(* IEC 61131-3 sources: JingjiangArm/moonboxpro_arm_8.4/Application/Application/数据类型/通讯协议/云影/读写内容/附属内容, 7 files *)

(* ---- StWrRd_AxisCfg.st ---- *)
(*@CES
Name=StWrRd_AxisCfg
Type=Gvl
TypeGuid=2db5746d-d284-4425-9f7f-2663a34b0ebc
Guid=0dd870ae-2077-401c-9916-294cbac50220
HasDeclaration=True
HasImplementation=False
*)
{DECLARATION}
{attribute 'pack_mode' := '1'}//系统配置
TYPE StWrRd_AxisCfg :
STRUCT
	xAxisProf_Enable: BIT;(*轴打开*)
	xAxisProf_MotRev: BIT;(*运动反向*)
	xAxisProf_SamRev: BIT;(*采样方向*)
	xAxisProf_Rsv1: BIT;(*预留*)
	xAxisProf_Rsv2: BIT;(*预留*)
	xAxisProf_Rsv3: BIT;(*预留*)
	xAxisProf_Rsv4: BIT;(*预留*)
	xAxisProf_Rsv5: BIT;(*预留*)

	//2025.11.1.104728两个字节作为站号通讯
	iSid: INT;
//	abyRsv: ARRAY [1..2] OF BYTE;(*预留两个字节方便增加其他内容*)
END_STRUCT
END_TYPE

{IMPLEMENTATION}

(* ---- StWrRd_MechanicalType.st ---- *)
(*@CES
Name=StWrRd_MechanicalType
Type=Gvl
TypeGuid=2db5746d-d284-4425-9f7f-2663a34b0ebc
Guid=03e174c8-9f43-4388-8870-9d21820ee6bb
HasDeclaration=True
HasImplementation=False
*)
{DECLARATION}
{attribute 'pack_mode' := '1'}
TYPE StWrRd_MechanicalType :
STRUCT
	byMachanicalTypeId: BYTE;(*1摆臂2直压3PVC直压4等料长5力达欧诺直压*)
	abyrsv: ARRAY [1..19] OF BYTE;//先放19个字节在这里放其他预套准相关内容|例如按钮
	abyBuffMechanicalParam: ARRAY [1..200] OF BYTE;(*机械参数*)
	//预留200字节用于通讯机械参数，
		//根据byMachanicalTypeId变量切换通讯内容
		//StMechanicalParam_01/
		//StMechanicalParam_02/
		//StMechanicalParam_03/
		//StMechanicalParam_05
END_STRUCT
END_TYPE

{IMPLEMENTATION}

(* ---- StWrRd_Switch_Grp.st ---- *)
(*@CES
Name=StWrRd_Switch_Grp
Type=Gvl
TypeGuid=2db5746d-d284-4425-9f7f-2663a34b0ebc
Guid=4a26eb77-6c13-4193-b710-63a532b0c18f
HasDeclaration=True
HasImplementation=False
*)
{DECLARATION}
{attribute 'pack_mode' := '1'}//总22字节
TYPE StWrRd_Switch_Grp :
STRUCT
	xSwitch_MachineRev							: BIT;(*反向走料开关*)
	xSwitch_6Inch_Rw							: BIT;(*收料3/6吋选择开关*)
	xSwitch_StartUp								: BIT;(*一键开机开关*)
	xSwitch_DiamMeasureAuto						: BIT;(*自动卷径开关*)
	xSwitch_RollOver							: BIT;(*设备翻料架开关*)
	xSwitch_Thickness							: BIT;(*料膜厚度手自动获取开关*)
	xSwitch_CutDneResetPidEn_Uw					: BIT;(*放料裁切后系数手自动*)
	xSwitch_CutDneResetPidEn_Rw					: BIT;(*收料裁切后系数手自动*)
	xSwitch_AutomaticCutEn_Uw					: BIT;(*放料自动接料是能*)
	xSwitch_AutomaticCutEn_Rw					: BIT;(*放料自动接料是能*)
	xSwitch_AutoAdjust_V_Grp					: BIT;(*整机纵向自动调整开关*)
	xSwitch_AutoAdjust_H_Grp					: BIT;(*整机纵向自动调整开关*)
	xSwitch_Follow_1U_V_Grp						: BIT;(*纵向跟1色开关*)
	xSwitch_Follow_1U_H_Grp						: BIT;(*横向跟1色开关*)
	xSwitch_DiamAuto_Pot						: BIT;(*卷径检测使用电位器*)
	xSwitch_DiamAuto_Enc						: BIT;(*卷径检测使用编码器*)
	xSwitch_DiamAuto_Ultrasonic_S				: BIT;(*卷径检测使用单超声波*)
	xSwitch_DiamAuto_Ultrasonic_D				: BIT;(*卷径检测使用双超声波*)
	xSwitch_DiamAuto_DualParam					: BIT;(*卷径检测双轴参数分开*)
	xSwitch_DebugMode							: BIT;(*调试模式开关*)
	xSwitch_Debug_DiamMeasure_Uw				: BIT;(*放料卷径检测电位器调试开关*)
	xBtn_Diameasure_Confirm_1					: BIT;(*自动卷径标定——1*)
	xBtn_Diameasure_Confirm_2					: BIT;(*自动卷径标定——2*)
	xBtn_Diameasure_Confirm_3					: BIT;(*自动卷径标定——3*)
	xBtn_Diameasure_Confirm_4					: BIT;(*自动卷径标定——4*)
(*2025.11.3.153321收放料绝对值编码器定位等相关开关
原总共42BIT位||重新整理一部分||总共需要14BIT位剩余作为预留*)
	xSwitch_UseAbsEnc_Uw						: BIT;(*放料使用绝对值编码器开关*)
	xSwitch_AxisLocaltion_DualParam_Uw			: BIT;(*放料绝对值编码器定位双轴参数开关*)
	xSwitch_Debug_Axis_Uw						: BIT;(*放料轴运行调试模式*)
	xSwitch_Debug_Uw_CutUpChoose				: BIT;(*放料绝对值编码器定位调试-上下裁选择||TRUE：上裁FALSE：下裁*)
	xSwitch_Debug_Uw_AxisA_Choose				: BIT;(*放料绝对值编码器定位调试-AB轴选择|TRUE:A轴；FALSE:B轴*)
	xBtn_Debug_Uw_Wr							: BIT;(*放料轴定位写入*)
	xBtn_Debug_Uw_MinDiam_Wr					: BIT;(*放料最小径写入*)
	xSwitch_UseAbsEnc_Rw						: BIT;(*收料使用绝对值编码器开关*)
	xSwitch_AxisLocaltion_DualParam_Rw			: BIT;(*收料绝对值编码器定位双轴参数开关*)
	xSwitch_Debug_Axis_Rw						: BIT;(*收料轴运行调试模式*)
	xSwitch_Debug_Rw_CutUpChoose				: BIT;(*收料绝对值编码器定位调试-上下裁选择||TRUE：上裁FALSE：下裁*)
	xSwitch_Debug_Rw_AxisA_Choose				: BIT;(*收料绝对值编码器定位调试-AB轴选择|TRUE:A轴；FALSE:B轴*)
	xSwitch_Debug_Rw_Inch3_CutUpChoose			: BIT;(*收料绝对值编码器定位调试-3/6吋选择|TRUE:3吋；FALSE:6吋*)
	xBtn_Debug_Rw_Wr							: BIT;(*收料轴定位写入*)
//2026.4.25.140018合并结构体|niu.j|增加5个变量
	xSwitch_StartAutoFind	: BIT;(*全自动套印开关*)
	xSwitch_EnFastPress		: BIT;(*当前色找到就合压使能*)
	xSwitch_SaveRS2File		: BIT;(*粗采样保存*)
	xSwitch_RFailure		: BIT;(*全自动套印粗采样失败校准*)
	xSwitch_FFailure		: BIT;(*全自动套印精采样失败校准按钮*)
// 	xRsv_Grp_1									: BIT;
// 	xRsv_Grp_2									: BIT;
// 	xRsv_Grp_3									: BIT;
// 	xRsv_Grp_4									: BIT;
// 	xRsv_Grp_5									: BIT;
//2026.4.25.140311增加结束
	xRsv_Grp_6									: BIT;
	xRsv_Grp_7									: BIT;
	xRsv_Grp_8									: BIT;
	xRsv_Grp_9									: BIT;
	xRsv_Grp_10									: BIT;
	xRsv_Grp_11									: BIT;
	xRsv_Grp_12									: BIT;
	xRsv_Grp_13									: BIT;
	xRsv_Grp_14									: BIT;
	xRsv_Grp_15									: BIT;
	xRsv_Grp_16									: BIT;
	xRsv_Grp_17									: BIT;
	xRsv_Grp_18									: BIT;
//2026.4.28.104338增加异站虚拟码盘重新配置开关xRsv_Grp_19
//	xRsv_Grp_19									: BIT;
	xSwitch_ReSetEncCfg							: BIT;

//bit20和bit21替换为换卷完成放料和收料
// 	xRsv_Grp_20									: BIT;
// 	xRsv_Grp_21									: BIT;
	xBtn_ChangeFilmDn_Uw						: BIT;
	xBtn_ChangeFilmDn_Rw						: BIT;
//2026.04.10.180829结束
//2026.03.11.100402 | + | 使用Bit22作为压力电机自动合压开关
	xSwitch_PressureAuto_Up_Dn							: BIT;
	//xRsv_Grp_22									: BIT;
//2026.2.25.094558 | + | 使用Bit23作为天枢数据保存的开关
	xSwitch_SaveData_GNS						: BIT;
	//xRsv_Grp_23									: BIT;
//2026.02.01.112053 | + | 使用Bit24作为停机维持使能的开关
	xSwitch_KeepServoOn							: BIT;
	//xRsv_Grp_24									: BIT;
//2026.01.27.093334 | + | 使用Bit25和Bit26作为清除报警按钮和回零位的操作标志
	xSwitch_ClearSysAlarm						: BIT;
	xSwitch_BackToHome							: BIT;
// 	xRsv_Grp_25									: BIT;
// 	xRsv_Grp_26									: BIT;
//2026.1.5.151405增加用Bit27和bit28作为收牵压力传感器调整开关和带长调整基准（标准带长/首色带长）开关（暂时只有秦华用）
	xSwitch_TensionAdjust_QH					: BIT;
	xSwitch_PrnLenAdj_Follow_QH					: BIT;
//	xRsv_Grp_27									: BIT;
//	xRsv_Grp_28									: BIT;
(*
	xSwitch_UseAbsEnc_Uw						: BIT;(*放料使用绝对值编码器开关*)
	xSwitch_AxisLocaltion_DualParam_Uw			: BIT;(*放料绝对值编码器定位双轴参数开关*)
	xSwitch_Debug_Axis_Uw						: BIT;(*放料轴运行调试模式*)
	xSwitch_Debug_Uw_CutUpChoose				: BIT;(*放料绝对值编码器定位调试-上裁选择*)
	xSwitch_Debug_Uw_AxisA_CutUpChoose			: BIT;(*放料绝对值编码器定位调试-上裁A选择*)
	xBtn_Debug_Uw_AxisA_CutUpWr					: BIT;(*上裁A轴定位写入*)
	xBtn_Debug_Uw_MinDiamA_CutUpWr				: BIT;(*上裁A轴最小径写入*)
	xSwitch_Debug_Uw_AxisB_CutUpChoose			: BIT;(*放料绝对值编码器定位调试-上裁B选择*)
	xBtn_Debug_Uw_AxisB_CutUpWr					: BIT;(*上裁B轴定位写入*)
	xBtn_Debug_Uw_MinDiamB_CutUpWr				: BIT;(*上裁B轴最小径写入*)
	xSwitch_Debug_Uw_CutDnChoose				: BIT;(*放料绝对值编码器定位调试-下裁选择*)
	xSwitch_Debug_Uw_AxisA_CutDnChoose			: BIT;(*放料绝对值编码器定位调试-下裁A选择*)
	xBtn_Debug_Uw_AxisA_CutDnWr					: BIT;(*下裁A轴定位写入*)
	xBtn_Debug_Uw_MinDiamA_CutDnWr				: BIT;(*下裁A轴最小径写入*)
	xSwitch_Debug_Uw_AxisB_CutDnChoose			: BIT;(*放料绝对值编码器定位调试-下裁B选择*)
	xBtn_Debug_Uw_AxisB_CutDnWr					: BIT;(*下裁B轴定位写入*)
	xBtn_Debug_Uw_MinDiamB_CutDnWr				: BIT;(*下裁B轴最小径写入*)
	xSwitch_UseAbsEnc_Rw						: BIT;(*收料使用绝对值编码器开关*)
	xSwitch_AxisLocaltion_DualParam_Rw			: BIT;(*收料绝对值编码器定位双轴参数开关*)
	xSwitch_Debug_Axis_Rw						: BIT;(*收料轴运行调试模式*)
	xSwitch_Debug_Rw_CutUpChoose				: BIT;(*收料绝对值编码器定位调试-上裁选择*)
	xSwitch_Debug_Rw_Inch3_CutUpChoose			: BIT;(*收料绝对值编码器定位调试-上裁3吋选择*)
	xSwitch_Debug_Rw_AxisA_3_CutUpChoose		: BIT;(*收料绝对值编码器定位调试-上裁A选择*)
	xBtn_Debug_Rw_AxisA_3_CutUpWr				: BIT;(*上裁A轴定位写入*)
	xSwitch_Debug_Rw_AxisB_3_CutUpChoose		: BIT;(*收料绝对值编码器定位调试-上裁B选择*)
	xBtn_Debug_Rw_AxisB_3_CutUpWr				: BIT;(*上裁B轴定位写入*)
	xSwitch_Debug_Rw_Inch6_CutUpChoose			: BIT;(*收料绝对值编码器定位调试-上裁6吋选择*)
	xSwitch_Debug_Rw_AxisA_6_CutUpChoose		: BIT;(*收料绝对值编码器定位调试-上裁A选择*)
	xBtn_Debug_Rw_AxisA_6_CutUpWr				: BIT;(*上裁A轴定位写入*)
	xSwitch_Debug_Rw_AxisB_6_CutUpChoose		: BIT;(*收料绝对值编码器定位调试-上裁B选择*)
	xBtn_Debug_Rw_AxisB_6_CutUpWr				: BIT;(*上裁B轴定位写入*)
	xSwitch_Debug_Rw_CutDnChoose				: BIT;(*收料绝对值编码器定位调试-下裁选择*)
	xSwitch_Debug_Rw_Inch3_CutDnChoose			: BIT;(*收料绝对值编码器定位调试-下裁3吋选择*)
	xSwitch_Debug_Rw_AxisA_3_CutDnChoose		: BIT;(*收料绝对值编码器定位调试-下裁A选择*)
	xBtn_Debug_Rw_AxisA_3_CutDnWr				: BIT;(*下裁A轴定位写入*)
	xSwitch_Debug_Rw_AxisB_3_CutDnChoose		: BIT;(*收料绝对值编码器定位调试-下裁B选择*)
	xBtn_Debug_Rw_AxisB_3_CutDnWr				: BIT;(*下裁B轴定位写入*)
	xSwitch_Debug_Rw_Inch6_CutDnChoose			: BIT;(*收料绝对值编码器定位调试-下裁6吋选择*)
	xSwitch_Debug_Rw_AxisA_6_CutDnChoose		: BIT;(*收料绝对值编码器定位调试-下裁A选择*)
	xBtn_Debug_Rw_AxisA_6_CutDnWr				: BIT;(*下裁A轴定位写入*)
	xSwitch_Debug_Rw_AxisB_6_CutDnChoose		: BIT;(*收料绝对值编码器定位调试-下裁B选择*)
	xBtn_Debug_Rw_AxisB_6_CutDnWr				: BIT;(*下裁B轴定位写入*)
*)
	xSwitch_Scrap_Avoidance						: BIT;(*裁切让料头开关*)
	xSwitch_CCW_AfterCut_Uw						: BIT;(*放料裁切后反转轴开关*)
	xSwitch_CutUseReflectionSensor				: BIT;(*放料裁切使用弧面开关*)
	xSwitch_UseRadCompensate_Uw					: BIT;(*放料翻转架补偿开关*)
	xSwitch_TowerDir_Uw							: BIT;(*翻转架补偿方向取反开关*)
	xBtn_ConfirmRad0_Uw							: BIT;(*放料翻转架补偿0弧度确认按钮*)
(*2025.11.14.145213调试使能只需要一个
	xSwitch_Debug_SpdAxisA_Uw					: BIT;(*放料A轴速度调试模式开关*)
	xBtn_DebugSpdAxisA_Uw_MoveEn				: BIT;(*放料A轴运动使能*)
	xBtn_DebugSpdAxisA_Uw_AccEn					: BIT;(*放料A轴加速使能*)
	xSwitch_Debug_SpdAxisB_Uw					: BIT;(*放料B轴速度调试模式开关*)
	xBtn_DebugSpdAxisB_Uw_MoveEn				: BIT;(*放料B轴运动使能*)
	xBtn_DebugSpdAxisB_Uw_AccEn					: BIT;(*放料B轴加速使能*)
	xSwitch_Debug_SpdAxisA_Rw					: BIT;(*收料A轴速度调试模式开关*)
	xBtn_DebugSpdAxisA_Rw_MoveEn				: BIT;(*收料A轴运动使能*)
	xBtn_DebugSpdAxisA_Rw_AccEn					: BIT;(*收料A轴加速使能*)
	xSwitch_Debug_SpdAxisB_Rw					: BIT;(*收料B轴速度调试模式开关*)
	xBtn_DebugSpdAxisB_Rw_MoveEn				: BIT;(*收料B轴运动使能*)
	xBtn_DebugSpdAxisB_Rw_AccEn					: BIT;(*收料B轴加速使能*)
	*)
	xSwitch_Debug_Spd_Uw					: BIT;(*放料A轴速度调试模式开关*)
	xBtn_DebugSpdAxisA_Uw_MoveEn				: BIT;(*放料A轴运动使能*)
	xBtn_DebugSpdAxisA_Uw_AccEn					: BIT;(*放料A轴加速使能*)
	xSwitch_Rsv1					 				: BIT;(*2025.11.14.145252原收料B轴速度调试模式开关*)
	xBtn_DebugSpdAxisB_Uw_MoveEn				: BIT;(*放料B轴运动使能*)
	xBtn_DebugSpdAxisB_Uw_AccEn					: BIT;(*放料B轴加速使能*)
	xSwitch_Debug_Spd_Rw					: BIT;(*收料A轴速度调试模式开关*)
	xBtn_DebugSpdAxisA_Rw_MoveEn				: BIT;(*收料A轴运动使能*)
	xBtn_DebugSpdAxisA_Rw_AccEn					: BIT;(*收料A轴加速使能*)
	xSwitch_Rsv					 				: BIT;(*2025.11.14.145252原收料B轴速度调试模式开关*)
	xBtn_DebugSpdAxisB_Rw_MoveEn				: BIT;(*收料B轴运动使能*)
	xBtn_DebugSpdAxisB_Rw_AccEn					: BIT;(*收料B轴加速使能*)

	xSwitch_UseFollow_1U_V_UwCut				: BIT;(*裁切套色新方式开关*)
	xSwitch_TypeGetInitDiam						: BIT;(*收放料初始卷径获取方式*)
	xSwitch_Heating_I							: BIT;(*全部加热1档*)
	xSwitch_Heating_II							: BIT;(*全部加热1I档*)
	xSwitch_Heating_III							: BIT;(*全部加热1II档*)
	xSwitch_Heating_Close						: BIT;(*全部加热关闭*)
	xSwitch_Heating_Water						: BIT;(*全部水加热控制开关*)
	xSwitch_Heating_Elc							: BIT;(*全部电加热控制开关*)
	xBtn_CopySV_1U_To_Other						: BIT;(*复制1色设定温度到其他色组*)
	xBtn_Reset_TempCtlBlock						: BIT;(*重启温控模块按钮*)
	xBtn_AllExhAir_On							: BIT;(*排风总开*)
	xBtn_AllExhAir_Off							: BIT;(*排风总关*)
	xBtn_CopyExhFreq_1U_To_Other				: BIT;(*复制1色设定温度到其他色组*)
	xBtn_ExhAir_Reset							: BIT;(*排风总关*)
	/////////////////////////////////////////////////////////////////////////////////////////////
	//以上刚好99bit，再增加9字节+5bit吧预留
	(*增加14BIT-9905界面*)
	xPidType_If_New								: BIT;
	xPidType_Of_New                 			: BIT;
	xBtn_StepTest_V                 			: BIT;
	xUseDiam_LowPass_Rw             			: BIT;
	xTensionCompensateEn_Rw         			: BIT;
	xUseTime_b1_Rw                  			: BIT;
	xUseTime_Variaition_Rw          			: BIT;
	xUseIMatrix_rX_DARE_Rw          			: BIT;
	xTensionCompensateEn_RwCut      			: BIT;
	xUseDiam_LowPass_Uw             			: BIT;
	xTensionCompensateEn_Uw         			: BIT;
	xUseTime_b1_Uw                  			: BIT;
	xUseTime_Variaition_Uw          			: BIT;
	xUseIMatrix_rX_DARE_Uw          			: BIT;

(**占用两个BIT位-卷径估计开关|2025.8.20.163450|niu.j
	xRsv_Flag0											: BIT;
	xRsv_Flag1											: BIT;
	*)
	xSwitch_Estimate_Uw					: BIT;(*放料卷径估计开关*)
	xSwitch_Estimate_Rw					: BIT;(*收料卷径估计开关*)

	xSwitchTension_If											: BIT;
	xSwitchTension_Of											: BIT;
	xUseBtn_Linkage											: BIT;
	xSwitch_ScraperOn_Of										: BIT;

	xNegPolarity_Uw											: BIT;
	xNegPolarity_Rw											: BIT;
	xNegPolarity_If											: BIT;
	xNegPolarity_Of											: BIT;

//2025.10.14.105504bit0和1、2、3用做dwControlBits.30和.31
	xSwitch_TempFromEnc_PT1000_If							: BIT;
	xSwitch_MotorTemp_PT1000_NTC_If						: BIT;
	xSwitch_TempFromEnc_PT1000_Of							: BIT;
	xSwitch_MotorTemp_PT1000_NTC_Of						: BIT;
//	xRsv_Flag0											: BIT;
//	xRsv_Flag1											: BIT;
//	xRsv_Flag2											: BIT;
//	xRsv_Flag3											: BIT;
//2025.10.14.111349|用bit4替代为xTensionCompensateEn_UwCut
	xTensionCompensateEn_UwCut							: BIT;
//	xRsv_Flag4											: BIT;
//2025.10.14.112844重新取出来一个byte用做位|bit0用作xUseAntiNotch_Uw
	xUseAntiNotch_Uw										: BIT;(*套色使用陷波器@*)
//2025.10.14.113357用bit1替代	xWorkMode_RollerPress					: BOOL;(*压辊顺序; TRUE从前到后; FALSE从后到前|*)
	xWorkMode_RollerPress										: BIT;
//	xRsv_Flag1										: BIT;
//2025.10.14.135539|用bit2和bit3替代等料长
	xSwitch_WaitFilmLengthEn				: BIT;(*开机等料长|原原wCtlSwitchRef.4*)
	xSwitch_WaitFilmLengthEn_From1st		: BIT;(*开机等首色料长|原原wCtlSwitchRef.13*)

//	xRsv_Flag2										: BIT;
//	xRsv_Flag3										: BIT;
//2025.10.15.144413|bit4用于套色报警铃
	xSwitch_Alarm_Arc						: BIT;(*套色报警开关|wCtlSwitchRef.0*)

//	xRsv_Flag4										: BIT;
//2025.10.15.160851||bit5和bit6用作预热风和预加热界面使能开关
	xSwitch_PreHotAirEn								: BIT;
	xSwitch_PreHeatingEn							: BIT;
//	xRsv_Flag5										: BIT;
//	xRsv_Flag6										: BIT;
//2025.10.15.165123||bit7和新的bi0-bit3用作刮刀递墨总控-再取一个BYTE用做BIT||5-1=4
	xSwitch_ScraperAuto					: BIT;(*刮刀手自动*)
	xSwitch_ScraperOn					: BIT;(*刮刀开关*)
	xSwitch_InkRollerAuto				: BIT;(*递墨辊手自动*)
	xSwitch_InkRollerCW					: BIT;(*递墨辊正转*)
	xSwitch_InkRollerCCW				: BIT;(*递墨辊反转*)
//	xRsv_Flag7										: BIT;
//	xRsv_Flag0										: BIT;
//	xRsv_Flag1										: BIT;
//	xRsv_Flag2										: BIT;
//	xRsv_Flag3										: BIT;
//2025.10.20.153333||bit4-bit7用做预套准按钮
	xBtn_ReadPhase_Home: BIT;//读取装版相位按钮
	xBtn_PreRegisterAxisId_Manu					: BIT;(*预套准的轴号手动确定@不考虑联动开关*)
	xBtn_PreRegister: BIT;//预套准按钮
	xBtn_PreRegisterCorrConfirm: BIT;//预套准自动修正按钮

	//xRsv_Flag4										: BIT;
	//xRsv_Flag5										: BIT;
	//xRsv_Flag6										: BIT;
	//xRsv_Flag7										: BIT;
	//再取一个BYTE用做BIT||4-1=3
	//2025.10.20.153729||bit0和bit1用作横向预套准按钮
	xBtn_HorzPreRegister_Repeat				: BIT;(*横向重复值按钮*)
	xBtn_HorzPreRegister_Setup				: BIT;(*横向设定值按钮*)

	//xRsv_Flag0										: BIT;
	//xRsv_Flag1										: BIT;
//2025.10.20.163844用bit2作为配方通讯标志
//金刚读取配方完成后，给天枢一个相位回复标志，天枢读取配方回复内容并且进行相位回复
	xBtn_RestorePhase_Hmi					: BIT;
//	xRsv_Flag2										: BIT;
//2025.12.30.171854||bit3和bit4用作界面切换上下裁开关
	xSwitch_Change_CutterOnTop_HMI_Uw				: BIT;
	xSwitch_Change_CutterOnTop_HMI_Rw				: BIT;
//	xRsv_Flag3										: BIT;
//	xRsv_Flag4										: BIT;
//2025.12.30.172757||bit5和bit6分别做收料3/6吋切换使用界面/开关，以及界面切换3/6吋开关
	xUseKnob_6Inch_Rw_Hmi							: BIT;
	xKnob_6Inch_Rw									: BIT;
//	xRsv_Flag5										: BIT;
//	xRsv_Flag6										: BIT;
//	xRsv_Flag7										: BIT;
	xSwitch_GrpInkEn:									BIT;
//2026.5.14.151101再取一位
	xSwitch_En_AutoStop								: BIT;
//xRsv_Flag1用作界面自动加减速按钮
	xAutoAccDec_Hmi									: BIT;
//	xRsv_Flag1										: BIT;

//2026.05.24.134141 增加光纤行走相关开关
//	xRsv_Flag2										:BIT;
// 	xRsv_Flag3										: BIT;
//	xRsv_Flag4										: BIT;
// 	xRsv_Flag5										: BIT;
// 	xRsv_Flag6										: BIT;
// 	xRsv_Flag7										: BIT;
	xFiberMove_DebugMode							:BIT;(*光纤行走调试模式*)
	xFiberMoveDisRunStart_AllUnit					:BIT;(*光纤行走同步运动启动*)
	xUseOnline_FiberMove							:BIT;(*光纤行走使用外部联动*)
	xFiberMoveConfirm_AllUnit						:BIT;(*光纤行走主站确认基准位置*)
	xFiberMovePosCal_ByUnit							:BIT;(*光纤行走色组标定*)
	xFiberMovePosCal_ByOnline						:BIT;(*光纤行走在线标定*)

	xFiberMove_Negative_AdjustByUnit				:BIT;(*光纤行走色组修正取反*)
	xFiberMove_Negative_AdjustByOnline				:BIT;(*光纤行走在线修正取反*)
	xRsv_Flag0										: BIT;
	xRsv_Flag1										: BIT;
	xRsv_Flag2										: BIT;
	xRsv_Flag3										: BIT;
	xRsv_Flag4										: BIT;
	xRsv_Flag5										: BIT;

	abyRsv_Flag											: ARRAY [1..1] OF BYTE;

END_STRUCT
END_TYPE

{IMPLEMENTATION}

(* ---- StWrRd_Switch_Machine.st ---- *)
(*@CES
Name=StWrRd_Switch_Machine
Type=Gvl
TypeGuid=2db5746d-d284-4425-9f7f-2663a34b0ebc
Guid=365f591a-c508-4b2d-a584-49adde6311bf
HasDeclaration=True
HasImplementation=False
*)
{DECLARATION}
TYPE StWrRd_Switch_Machine ://总12字节
STRUCT
	xSwitch_PreHotEn_Print								: BIT;(*预热印刷激活开关*)
	xSwitch_ExhAir_Limit_HotWind						: BIT;(*排风限制热风开关*)
	xSwitch_ExhAir_Limit_Run							: BIT;(*排风限制开机开关*)
	xSwitch_CommEn_WatchDevice_Tcp						: BIT;(*TCP-外部监控设备开关*)
	xSwitch_CommEn_WatchDevice_485						: BIT;(*485-外部监控设备开关*)
	xSwitch_CommEn_1U_485								: BIT;(*1色人机通讯开关*)
	xSwitch_CommEn_485									: BIT;(*485通讯开关*)
	xSwitch_CommEn_485_Exh								: BIT;(*排风485通讯开关*)
	xSwitch_CommEn_485_Scraper							: BIT;(*刮刀485通讯开关*)
	xSwitch_CommEn_485_InkRoller						: BIT;(*递墨辊485通讯开关*)
	xSwitch_CommEn_485_HotWind							: BIT;(*热风485通讯开关*)
	xSwitch_ArcIntensityBtn_Hmi							: BIT;(*手动调节随速度走开关*)
	xSwitch_PrnRatioIndividual_Setting					: BIT;(*色组版辊减速比单独设置开关*)
	xSwitch_NetRatioIndividual_Setting					: BIT;(*色组网辊减速比单独设置开关*)
	xSwitch_BottomRatioIndividual_Setting				: BIT;(*色组底辊减速比单独设置开关*)
	xSwitch_StepDriveDebugRun							: BIT;(*横向步进电机测试执行开关*)
	/////////////////////////////////////////////////////////////////////////////////////////////
	//以上刚好16bit，再增加10字节吧预留
	//增加21BIT
	xSetProPointEn										: BIT;
	xUseMaxTimeAsSBegin_InLowSpeed      				: BIT;
	xPseudoRandomEn                     				: BIT;
	xPseudoRandomStart                  				: BIT;
	xEn_RevLimit                        				: BIT;
	xSaveFineSampleData_ToArc           				: BIT;
	xReqSetLedFunc                      				: BIT;
	xSetHmiResolution                   				: BIT;
	xPopupWindowVisible                 				: BIT;
	xInitArcErr_AjdImmediately          				: BIT;
	xPhaseAutoRecoveryEn                				: BIT;
	xKeepServo_PreRegisterDne           				: BIT;
	xUseIfVel_Uw                        				: BIT;
	xKeepServo_Stop                     				: BIT;
	xAxisPrfVelEn                       				: BIT;
	xUseGc_PID_2025                     				: BIT;
	xFlag_Follow_1U_Double_V            				: BIT;
	xArcErrCorrectIsRev_V               				: BIT;
	xAutoSetSampleType                  				: BIT;
	xGetSampleTypeBtn                   				: BIT;
	xAutoSetArcCtlWay                   				: BIT;

	xWorkMode_Inch										: BIT;

//bit1和bit2代替为g_xScraperReset和g_xInkRollerReset
	xSwitch_ScraperReset								: BIT;
	xSwitch_InkRollerReset								: BIT;
//	xRsv_Flag1											: BIT;
//	xRsv_Flag2											: BIT;
//2025.10.14.145403取一个BYTE当做BIT位处理7-1=6
	xSwitch_HotwindReset: BIT;
	xSwitch_ResetTemctlModule: BIT;
	xMoveFreq_I_ToAll_AirHot: BIT;
	xMoveFreq_II_ToAll_AirHot: BIT;
	xMoveFreq_III_ToAll_AirHot: BIT;
	xMoveFreq_I_ToAll_ExhaustAir: BIT;
	xMoveFreq_II_ToAll_ExhaustAir: BIT;
	xMoveFreq_III_ToAll_ExhaustAir: BIT;
//2025.10.14.151736取一个BYTE当用bit6-1=5
	xSwitch_Copy1stUExhaustDamperPos : BIT;
//2025.11.6.134235||bit1用来作为保存系统配置按钮通讯
	xBtn_UpdateSysCfg: BIT;
//	xBITrsv1: BIT;
//2026.1.5.150714||bit2/bit3用做底辊周长/减速比单独设定开关||bit4/bit5用做网辊周长/减速比单独设定开关
	xSwitch_IndependentSettings_BottomGirth: BIT;
	xSwitch_IndependentSettings_BottomRatio: BIT;
	xSwitch_IndependentSettings_NetGirth: BIT;
	xSwitch_IndependentSettings_NetRatio: BIT;

// 	xBITrsv2: BIT;
// 	xBITrsv3: BIT;
// 	xBITrsv4: BIT;
// 	xBITrsv5: BIT;
	xBITrsv6: BIT;
	xBITrsv7: BIT;

	abyRsv_Flag											: ARRAY [1..5] OF BYTE;

END_STRUCT
END_TYPE

{IMPLEMENTATION}

(* ---- StWrRd_Switch_Unit.st ---- *)
(*@CES
Name=StWrRd_Switch_Unit
Type=Gvl
TypeGuid=2db5746d-d284-4425-9f7f-2663a34b0ebc
Guid=a2047d0e-672b-403c-b194-95cddde93ad4
HasDeclaration=True
HasImplementation=False
*)
{DECLARATION}
{attribute 'pack_mode' := '1'}//总16字节
TYPE StWrRd_Switch_Unit :
STRUCT
	xSwitch_CoatingPrn					: BIT;(*色组涂布开关*)
	xSwitch_CoatingRec					: BIT;(*涂布调整反向*)
	xSwitch_ScraperAuto					: BIT;(*刮刀手自动*)
	xSwitch_ScraperOn					: BIT;(*刮刀开关*)
	xSwitch_InkRollerAuto				: BIT;(*递墨辊手自动*)
	xSwitch_InkRollerCW					: BIT;(*递墨辊正转*)
	xSwitch_InkRollerCCW				: BIT;(*递墨辊反转*)
	xSwitch_HotWindOn					: BIT;(*热风开关*)
	xSwitch_HeatingOn					: BIT;(*加热开关*)
	xSwitch_Heating_I					: BIT;(*加热I档*)
	xSwitch_Heating_II					: BIT;(*加热II档*)
	xSwitch_Heating_III					: BIT;(*加热III档*)
	xSwitch_ThisUnitEna					: BIT;(*色组套印开关*)
	xSwitch_Horz						: BIT;(*横向开关*)
	xSwitch_DoorBaseLn					: BIT;(*门内基线开关*)

	xSwitch_SmallSignalProcessing_T1	: BIT;(*第一组波门T1内小信号处理开关*)
	xSwitch_SmallSignalProcessing_T2	: BIT;(*第一组波门T2内小信号处理开关*)
	xSwitch_Rsv_1						: BIT;
	xSwitch_Rsv_2						: BIT;
(*	2025.10.27.141051||小信号只有两个T1和T2，不用分波门
	xSwitch_SmallSignalProcessing_T1_1	: BIT;(*第一组波门T1内小信号处理开关*)
	xSwitch_SmallSignalProcessing_T2_1	: BIT;(*第一组波门T2内小信号处理开关*)
	xSwitch_SmallSignalProcessing_T1_2	: BIT;(*第二组波门T1内小信号处理开关*)
	xSwitch_SmallSignalProcessing_T2_2	: BIT;(*第二组波门T2内小信号处理开关*)
	*)
	xSwitch_AutoAdjust_V_Unit			: BIT;(*整机纵向自动调整开关*)
	xSwitch_AutoAdjust_H_Unit			: BIT;(*整机纵向自动调整开关*)
	xSwitch_NegativePolarity_T1_1		: BIT;(*第一组波门内T1信号反极性*)
	xSwitch_NegativePolarity_T2_1		: BIT;(*第一组波门内T2信号反极性*)
	xSwitch_NegativePolarity_T1_2		: BIT;(*第二组波门内T1信号反极性*)
	xSwitch_NegativePolarity_T2_2		: BIT;(*第二组波门内T2信号反极性*)
	xSwitch_AdjRev_V					: BIT;(*纵向调整反*)
	xSwitch_AdjRev_H					: BIT;(*横向调整反*)
	xSwitch_AdjRev_O					: BIT;(*单标记调整反*)
	xSwitch_Follow_1U_V_Unit			: BIT;(*纵向跟1色开关*)
	xSwitch_Follow_1U_H_Unit			: BIT;(*横向跟1色开关*)
	xSwitch_DualPolarity				: BIT;(*双极性开关*)
	xSwitch_UnitRevPrn					: BIT;(*色组反印开关*)
	xSwitch_DualGate					: BIT;(*双波门开关*)
	xSwitch_Transfer_Err				: BIT;(*误差传递开关*)
	xSwitch_Transfer_Adj				: BIT;(*调整量传递开关*)
(*卷径估计与色组无关|2025.8.20.163318|niu.j|放出两个BIT位
	xSwitch_Estimate_Uw					: BIT;(*放料卷径估计开关*)
	xSwitch_Estimate_Rw					: BIT;(*收料卷径估计开关*)
	*)
//占用xRsv_Flag1作为印长调整开关2025.12.31.112738
	xSwitch_AdjBandLen					: BIT;
//	xRsv_Flag1							: BIT;
	xRsv_Flag2							: BIT;

	xSwitch_Heating_Water				: BIT;(*水加热控制开关*)
	xSwitch_Heating_Elc					: BIT;(*电加热控制开关*)
	xSwitch_ExhAir						: BIT;(*色组排风开关*)

	/////////////////////////////////////////////////////////////////////////////////////////////
	//以上刚好40bit，再增加11字节吧预留
	//2025.7.3.175755增加7BIT
	xCompensateEn_H						: BIT;
	xUseAntiNotch_Arc   				: BIT;
	xUsePeriodic    					: BIT;
	T1_S         						: BIT;
	T2_S         						: BIT;
	PT1000_M    						: BIT;
	ENCTMP_M     						: BIT;
	xSwitch_HorzMoveLeft_Manu_1							: BIT;(*横向左调0.01*)
	xSwitch_HorzMoveLeft_Manu_2							: BIT;(*横向左调0.02*)
	xSwitch_HorzMoveLeft_Manu_3							: BIT;(*横向左调0.05*)
	xSwitch_HorzMoveRight_Manu_1						: BIT;(*横向右调0.01*)
	xSwitch_HorzMoveRight_Manu_2						: BIT;(*横向右调0.02*)
	xSwitch_HorzMoveRight_Manu_3						: BIT;(*横向右调0.05*)
//2025.10.14.105504bit6和7用做dwControlBits.30和.31
//	xRsv_Flag6											: BIT;
//	xRsv_Flag7											: BIT;
	xSwitch_TempFromEnc_PT1000							: BIT;
	xSwitch_MotorTemp_PT1000_NTC						: BIT;
//2025.12.30.222739变量xUnitExhaustDamperCtl_Auto占用Bit8||
	xUnitExhaustDamperCtl_Auto							: BIT;//排风风门控制自动
	//xRsv_Flag8											: BIT;
	(*2025.9.20.092456占用一个byte用于通讯界面横向手动按钮10-1=9*)

//2026.2.2.162623再取一个BYTE用做位处理2026.2.2.162710||niu.j||9-1=8
//取bit00用做清除标定按钮
	xSwitch_ResetFlag_FinishCalid						: BIT;
//	xRsv_Flag00											: BIT;
//取bit01用作标定模式界面开关
//	xSwitch_ModeCalib_Press								: BIT;
//	xRsv_Flag01											: BIT;
	xSwitch_Linkage										: BIT;//色组联动开关
	xSwitch_Ink											: BIT;//匀墨开关
//	xRsv_Flag02											: BIT;
//2026.4.24.144718||程序合并||新增6bit位||预留全部占完，需要新开一个byte
	xBtn_ConfirmLimit_Left								: BIT;//横向标定左
	xBtn_ConfirmLimit_Right								: BIT;//横向标定右
	xBtn_ResetLimit_Left								: BIT;//清除标定
	xBtn_ResetLimit_Right								: BIT;//清除标定
	xBtn_MoveLeft_Horz									: BIT;//横向左移
	xBtn_MoveRight_Horz									: BIT;//横向右移
//2026.4.24.145339结束
//2026.4.6.103029|占用两个变量处理全自动套印相关；bit3 he 4
	xSwitch_CurManuAdjust							: BIT;//(*当前色未找到，需要手动调整光电眼位置，调整好后人工置位*)
	xSwitch_PreCurManuAdjust						: BIT;//(*前一色未找到，需要观察原因调整好后，人工点确定，等一个机组料长后置位*)
//	xRsv_Flag00										    : BIT;
//	xRsv_Flag01											: BIT;
//本次占用结束2026.4.6.103323
//占用一个，做冷风开关
//	xRsv_Flag02											: BIT;
	xSwitch_CoolWind									: BIT;
//2026.5.29.171622结束
	xRsv_Flag03											: BIT;
	xRsv_Flag04									  		: BIT;
	xRsv_Flag05											: BIT;
	xRsv_Flag06											: BIT;
	abyRsv_Flag: ARRAY [1..7] OF BYTE;
END_STRUCT
END_TYPE

{IMPLEMENTATION}

(* ---- StWrRd_SysCfg.st ---- *)
(*@CES
Name=StWrRd_SysCfg
Type=Gvl
TypeGuid=2db5746d-d284-4425-9f7f-2663a34b0ebc
Guid=80b81a88-c08a-42a7-913a-d9e7c94af84c
HasDeclaration=True
HasImplementation=False
*)
{DECLARATION}
{attribute 'pack_mode' := '1'}//系统配置
TYPE StWrRd_SysCfg :
STRUCT
	iCompanyId					: INT := 0;(* 公司id/0科赛/1飞达/... *)
	byLanguageId				: BYTE := 1;(* 语言id/1.中文/2.英文/... *)
	byUnitMaxNum				: BYTE := 7;(* 色组数量/0~MAX_UNIT_NUM *)
	astStAxisCfgStruct_PC_		: ARRAY [1..MAX_UNIT_NUM] OF StWrRd_AxisCfg;(*光电眼行走机构 | 2024.04.01.092649*)
	astStAxisCfgStruct_BR_		: ARRAY [1..MAX_UNIT_NUM] OF StWrRd_AxisCfg;(* BR: Bottom Roller/底辊 *)
	astStAxisCfgStruct_PR_		: ARRAY [1..MAX_UNIT_NUM] OF StWrRd_AxisCfg;(* PR: Prn Roller/版辊 *)
	astStAxisCfgStruct_NR_		: ARRAY [1..MAX_UNIT_NUM] OF StWrRd_AxisCfg;(* NR: Net Roller/网辊 *)
	astStAxisCfgStruct_UW_I		: ARRAY [1..2] OF StWrRd_AxisCfg;(* UW: UnWind/放料 *)
	astStAxisCfgStruct_RW_I		: ARRAY [1..2] OF StWrRd_AxisCfg;(* RW: ReWind/收料 *)
	stStAxisCfgStruct_IF_I		: StWrRd_AxisCfg;(* IF: InFeed/放牵 *)
	stStAxisCfgStruct_OF_I		: StWrRd_AxisCfg;(* OF: OutFeed/收牵 *)
	astStAxisCfgStruct_CD_I		: ARRAY [1..2] OF StWrRd_AxisCfg;(* CD: Central Drum/中心滚筒 *)(*中心辊增加一个|2024.04.01.094732*)
(*以上总共220字节2025.10.13.104636*)

	astStAxisCfgStruct_PR_M_	: ARRAY [1..MAX_UNIT_NUM] OF StWrRd_AxisCfg;(* PR_M: PrnRoller Mside/版辊压力M侧 *)
	astStAxisCfgStruct_PR_G_	: ARRAY [1..MAX_UNIT_NUM] OF StWrRd_AxisCfg;(* PR_G: PrnRoller Gside/版辊压力G侧 *)
	astStAxisCfgStruct_NR_M_	: ARRAY [1..MAX_UNIT_NUM] OF StWrRd_AxisCfg;(* NR_M: NetRoller Mside/网辊压力M侧 *)
	astStAxisCfgStruct_NR_G_	: ARRAY [1..MAX_UNIT_NUM] OF StWrRd_AxisCfg;(* NR_G: NetRoller Gside/网辊压力G侧 *)
	astStAxisCfgStruct_UW_II		: ARRAY [1..2] OF StWrRd_AxisCfg;(* UW: UnWind/放料 *)
	astStAxisCfgStruct_RW_II		: ARRAY [1..2] OF StWrRd_AxisCfg;(* RW: ReWind/收料 *)
	stStAxisCfgStruct_IF_II		: StWrRd_AxisCfg;(* IF: InFeed/放牵 *)
	stStAxisCfgStruct_OF_II		: StWrRd_AxisCfg;(* OF: OutFeed/收牵 *)
	astStAxisCfgStruct_CD_II		: ARRAY [1..2] OF StWrRd_AxisCfg;(* CD: Central Drum/中心滚筒 *)(*中心辊增加一个|2024.04.01.094732*)
	abyDataRsv					: ARRAY [1..4] OF BYTE;
(*以上总共216+4字节2025.10.13.104657|*)

	astStAxisCfgStruct_STR_M_	: ARRAY [1..MAX_UNIT_NUM] OF StWrRd_AxisCfg;(* NR_M: NetRoller Mside/张带辊压力M侧 *)
	astStAxisCfgStruct_STR_G_	: ARRAY [1..MAX_UNIT_NUM] OF StWrRd_AxisCfg;(* NR_G: NetRoller Gside/张带辊压力G侧 *)
	astStAxisCfgStruct_HORIZ_	: ARRAY [1..MAX_UNIT_NUM] OF StWrRd_AxisCfg;(* HORIZ: 横向控制电机 *)
//	abyDataRsv1					: ARRAY [1..76] OF BYTE;
//2026.5.15.154633增加色组控制器配置|总48字节|76-48=28
	astStAxisCfgStruct_Ctl		: ARRAY [1..MAX_UNIT_NUM] OF StWrRd_AxisCfg;(*色组控制器配置通讯*)
	abyDataRsv1					: ARRAY [1..28] OF BYTE;
(*系统配置总共220*3个字节2025.10.13.105513*)
END_STRUCT
END_TYPE

{IMPLEMENTATION}

(* ---- StWrRd_UnitParam.st ---- *)
(*@CES
Name=StWrRd_UnitParam
Type=Gvl
TypeGuid=2db5746d-d284-4425-9f7f-2663a34b0ebc
Guid=921fa842-8dc1-46c6-9dca-e62db1c4c4c1
HasDeclaration=True
HasImplementation=False
*)
{DECLARATION}
{attribute 'pack_mode' := '1'}
TYPE StWrRd_UnitParam :
STRUCT
	stBitStWrRd_Switch_Unit							: StWrRd_Switch_Unit;(*总16*16字节*)
	rGirth_Using_CoatingPrn							: REAL;(*涂布周长*)
	byBtn_AdjModeSwitch_CoatingPrn					: BYTE;(*涂布调整方式切换按钮*)
	rStep_OfChangeGirth								: REAL;(*涂布版轴修改步幅*)
	rHz_UnitScraper_ManuallySet						: REAL;(*刮刀手动频率*)
	rCoeff_UnitScraper_Auto							: REAL;(*刮刀自动系数*)
	rHz_UnitInkRoller_ManuallySet					: REAL;(*递墨辊手动频率*)
	rCoeff_UnitInkRoller_Auto						: REAL;(*递墨辊自动系数*)
	rHz_UnitHotWind_ManuallySet						: REAL;(*热风手动频率*)
	rSV_UnitTemCtl									: REAL;(*加热设定温度*)
	iGateWidthPhy									: INT;(*波门宽度*)
	rAlarm_V										: REAL;(*纵向报警值*)
	rAlarm_H										: REAL;(*横向报警值*)
	rAdjust_V										: REAL;(*纵向修正量*)
	rAdjust_H										: REAL;(*横向修正量*)
	rDeadzoneMax_H									: REAL;(*横向最大不动作区*)
	rDeadzoneMin_H									: REAL;(*横向最小不动作区*)
	iCoefOfCoupling_V								: INT;(*纵向传递2系数*)
	byAverage_V										: BYTE;(*纵向平均值*)
	byAverage_H										: BYTE;(*横向平均值*)
	(*2025.8.20.161154|这里重新分配输出测试吧2025.8.20.161207|niu.j|先释放这里的空间*)
	(*awOutput_IOtestDO_Axis							: ARRAY [1..8] OF WORD;(*主面板IO测试输出*)
	awOutput_IOtestAO_Axis							: ARRAY [1..16] OF WORD;(*主面板IO测试输出*)*)

	(*2025.9.19.123648|niu.j|增加色组顺逆序选择|48-2=46*)
	iMarkArrangeMode							: INT;(* 标记排列方式 *)

//2025.10.20.151240||增加预套准相关参数|niu.j|46-10=36
	rPreReg_Adjust							: REAL;(*预套准调整量|*)
	rPreReg_ConstVal						: REAL;(*预套准色组间固定料长部分|单位:mm*)
	uiTurnOverFilmLenth						: UINT;(*翻料架料膜长度@mm*)
//2025.10.20.153028增加横向预套准参数36-12=24
	diPreReg_RepeatVal_H					: DINT;(*预套准重复值-横向|单位:mm|*)
	diPreReg_SetupVal_H						: DINT;(*预套准设定值-横向|单位:mm|*)
	diPreReg_AdjustVal_H					: DINT;(*预套准修正值*)

//2025.10.23.104815||增加一些配方里需要保存的内容24-14=10
	rGirth_PrnRoller					: REAL;
	iMarkTypeId_Pu						: INT;
	byAirInletWindDoorValue				: BYTE;
	byOvensAirOutWindDoorValue			: BYTE;
	byAirExhaustWindDoorValue			: BYTE;
	byAirReturnWindDoorValue			: BYTE;
	rHz_UnitHotWind_2_ManuallySet		: REAL;

//2025.12.30.223020|增加排风风门位置手动设定值||10-4=6
	rUnitExhaustDamperPos_ManuallySet		: REAL;(*排风风门位置手动设置值*)
//2025.12.31.112556增加带长调整一些参数|2字节|6-2=4
	iBandLengthFilterCnt					: INT;//带长滤波次数
	abyRsvData_2										: ARRAY [1..4] OF BYTE;

	uiTimeMs_RollerPressUpKeep						: UINT;(*压辊双气缸-离压保持时间*)
	uiAxisNum										: UINT;(*色组单独减速比分子*)
	uiAxisDen										: UINT;(*色组单独减速比分母*)
	rHz_UnitExhaust_ManuallySet						: REAL;(*色组排风设定频率*)

//9905界面内容

	rAxisVelPrf_Coeff1								: REAL;
	rAxisVelPrf_Coeff2             					: REAL;
	rAxisVelPrf_Coeff3             					: REAL;
	rMargin_Mag_Arc                					: REAL;
	//2026.05.13.091818+变量替换
	//rMargin_Phi_Arc                					: REAL;
	rKadj_I_Mol                					: REAL;
//	rMargin_Phi_Arc                					: REAL;
//2026.5.13.144804
//2026.4.25.142452结束
///	rKp_MolCal                     					: REAL;
///	rKi_MolCal                     					: REAL;
	abyRsv_Data_2									: ARRAY [1..8] OF BYTE;
//2026.4.25.142452结束
	rFilmLengthFromPrevPressUnit   					: REAL;
	byCompensateValue_Hor							: BYTE;
	byMaxAddValue_Total_Hor							: BYTE;
	rWn_Arc											: REAL;
	rBw_Arc											: REAL;
	rDp_Arc											: REAL;
	rK     											: REAL;
	rA2    											: REAL;
	rA1    											: REAL;
	rA0    											: REAL;
	rG_Periodic  									: REAL;
	rW_Periodic  									: REAL;
	byCnt_Comm2ARM									: BYTE;

//2025.7.3.175755以上总共208字节
////////////////////////////////////////////////////////////分割线///////////////////////////////////////////////
	(*增加一个波门位置2025.8.25.151314*)
	iGateSa											: INT;
	iGateSaEx										: INT;
//2025.10.20.142338增加纵横向飞点阈值|8-2=6
	byFakeThreshold_V				:BYTE;(*纵向飞点阀值@丝			*)
	byFakeThreshold_H				:BYTE;(*横向飞点阀值@丝			*)
//2025.10.20.143054增加界面显示误差平均次数6-1=5
	byAve_v_extra							: BYTE;(*界面误差显示平均值*)

	abyRsvData_0										: ARRAY [1..5] OF BYTE;

/////////////////////////////////////////////////////2025.7.3.175755新增12字节，总大小220byte//////////////////////////////////////////////////////////////
	abyRsvData_1										: ARRAY [1..440] OF BYTE;
	//2025.8.20.161050|niu.j|增加色组输出测试
	awOutput_IOtestDO_Axis							: ARRAY [1..4] OF WORD;(*主面板IO测试输出*)
	awOutput_IOtestAO_Axis							: ARRAY [1..6] OF WORD;(*主面板IO测试输出*)
	awOutput_IOtestDO_Axis_Extra					: ARRAY [1..6] OF WORD;(*主面板IO测试输出*)
	awOutput_IOtestAO_Axis_Extra					: ARRAY [1..24] OF WORD;(*主面板IO测试输出*)
//2026.1.5.175104||增加一些变量总共16字节，140-16=124
	rGirth_BottomGirth								: REAL;
	rGirth_NetGirth									: REAL;
	uiNum_Bottom									: UINT;
	uiDen_Bottom									: UINT;
	uiNum_Net										: UINT;
	uiDen_Net										: UINT;
	//2026.2.2.161811增加界面的一些开关|niu.j|总4*3个字节12||124-12=112
	adwPressureMotor_Move_MasterHMI					: ARRAY [1..3] OF DWORD;
	//2026.04.02.191022 增加横向限位实时位置|Hou.N|112-12=100
 	diPos_LimitLeft									:DINT;
 	diPos_LimitRight								:DINT;

	abyData_rsv_h									: ARRAY [1..4] OF BYTE;
 	//diPos_Horz										:DINT;
	//2026.05.24.135408增加光纤行走变量|xi.hy|100-12=88
	rFiberMoveAdjust								:REAL;(*光纤行走色组修正量*)
	rFiberMoveAdjust_ByOnlie						:REAL;(*光纤行走在线修正量*)
	uiFiberMove_SoftLimit_Min						:UINT;(*光纤行走左限位*)
	uiFiberMove_SoftLimit_Max						:UINT;(*光纤行走右限位*)

	//2026.5.29.172149增加金刚火眼误差/月光宝盒误差获取与调整选择||88-1=87
	byGetErrMode									: BYTE;
	//2026.06.15.183819 增加电压设定值 0-220V | 87-3=84
	abyVoltage_SV:ARRAY [1..3] OF BYTE;
	abyRsvData_3									: ARRAY [1..84] OF BYTE;

//	abyRsvData_3									: ARRAY [1..100] OF BYTE;
END_STRUCT
END_TYPE

{IMPLEMENTATION}
